(* IEC 61131-3 sources: P26002_Bosch_HDPump/P26002_Bosch_HDPump_PLC/RPM_Profiles, 4 files *)

(* ---- FB_ArrayProfile.st ---- *)
(********************************************************************************
 * FUNCTION_BLOCK: FB_ArrayProfile
 *
 * Beschreibung:
 *   Liest ein 10-ms-Raster Drehzahlprofil aus dem globalen Array aLapData
 *   und interpoliert im 1-ms-Takt stufenlos linear.
 *   Bei Erreichen von nPointsInLap springt der Zeiger auf 0 zurück und
 *   bLapFinished wird für einen Zyklus TRUE.
 ********************************************************************************)
FUNCTION_BLOCK FB_ArrayProfile
VAR_INPUT
    bExecute        : BOOL;
    nPointsInLap    : DINT; (* Tatsächliche Anzahl Punkte im Zyklus *)
END_VAR
VAR_IN_OUT
    aLapDataBuffer  : ARRAY[0..179999] OF REAL; (* Referenz auf das Daten-Array *)
END_VAR
VAR_OUTPUT
    fRpmOut         : REAL;
    bLapFinished    : BOOL;
END_VAR
VAR
    nIndex          : DINT := 0;
    nSubStep1ms     : INT  := 0;
    fCurrentP       : REAL;
    fNextP          : REAL;
    fDeltaPerMs     : REAL;
END_VAR

bLapFinished := FALSE;

(* Plausibilitätsprüfung *)
IF NOT bExecute OR (nPointsInLap <= 1) OR (nPointsInLap > 180000) THEN
    nIndex       := 0;
    nSubStep1ms  := 0;
    fRpmOut      := 0.0;
    RETURN;
END_IF;

(* Alle 10 ms: Neuer Stützwert aus dem Array *)
IF nSubStep1ms = 0 THEN
    fCurrentP := aLapDataBuffer[nIndex];

    (* Nächsten Punkt für Steigungsberechnung holen *)
    IF (nIndex + 1) < nPointsInLap THEN
        fNextP := aLapDataBuffer[nIndex + 1];
    ELSE
        fNextP := aLapDataBuffer[0]; (* Zyklischer Sprung zum Anfang *)
    END_IF;

    (* Steigung pro 1 ms berechnen *)
    fDeltaPerMs := (fNextP - fCurrentP) / 10.0;

    nIndex := nIndex + 1;

    (* RUNDENENDE: Letzter Punkt des Profils erreicht *)
    IF nIndex >= nPointsInLap THEN
        nIndex       := 0;    (* Für nächste Runde zurücksetzen *)
        bLapFinished := TRUE; (* Lap-Signal auslösen *)
    END_IF;
END_IF;

(* 1-ms-Interpolation *)
fRpmOut := fCurrentP + (fDeltaPerMs * INT_TO_REAL(nSubStep1ms));

(* 1-ms-Zähler 0 bis 9 *)
nSubStep1ms := (nSubStep1ms + 1) MOD 10;

END_FUNCTION_BLOCK

(* ---- FB_SequenceController.st ---- *)
(********************************************************************************
 * FUNCTION_BLOCK: FB_SequenceController
 *
 * Beschreibung:
 *   Steuert den Gesamt-Ablauf (Start/Stop, Wiederholungen, Gesamtdauer).
 *   Ausgänge:
 *     - bSequenceActive: TRUE ab Start bis zum Ende der gesamten Sequenz
 *     - bLapTrigger:     Gepulster Ausgang (z.B. 50ms) nach jedem Lap-Durchlauf
 ********************************************************************************)
FUNCTION_BLOCK FB_SequenceController
VAR_INPUT
    bStart              : BOOL;
    bStop               : BOOL;
    eEndMode            : E_SequenceEndMode;
    nTargetLaps         : UDINT;
    tTargetDuration     : TIME;
    tLapPulseDuration   : TIME := T#50ms; (* Einstellbare Pulsdauer *)
    bLapFinishedSignal  : BOOL;
    tCycleTime          : TIME := T#1ms;
END_VAR
VAR_OUTPUT
    bSequenceActive     : BOOL; (* Start/End-Trigger *)
    bLapTrigger         : BOOL; (* Gepulster Lap-Trigger *)
    nCompletedLaps      : UDINT;
    tElapsedTime        : TIME;
END_VAR
VAR
    bStartOld           : BOOL;
    nPulseCyclesLeft    : DINT := 0; (* Exakter Zyklustimer für den Puls *)
END_VAR

(* Stop-Befehl *)
IF bStop THEN
    bSequenceActive  := FALSE;
    nPulseCyclesLeft := 0;
END_IF;

(* Start-Flanke *)
IF bStart AND NOT bStartOld AND NOT bSequenceActive THEN
    bSequenceActive  := TRUE;
    nCompletedLaps   := 0;
    tElapsedTime     := T#0s;
    nPulseCyclesLeft := 0;
END_IF;
bStartOld := bStart;

(* Sequenz-Ablauf *)
IF bSequenceActive THEN
    tElapsedTime := tElapsedTime + tCycleTime;

    (* Lap-Ende registriert *)
    IF bLapFinishedSignal THEN
        nCompletedLaps   := nCompletedLaps + 1;
        (* Millisekunden in 1ms-Taskzyklen konvertieren *)
        nPulseCyclesLeft := TIME_TO_DINT(tLapPulseDuration);
    END_IF;

    (* Abbruchbedingungen *)
    CASE eEndMode OF
        MODE_LAP_COUNT:
            IF nCompletedLaps >= nTargetLaps THEN
                bSequenceActive := FALSE;
            END_IF;

        MODE_TIME_LIMIT:
            IF tElapsedTime >= tTargetDuration THEN
                bSequenceActive := FALSE;
            END_IF;
    END_CASE;
END_IF;

(* Deterministischer Puls über Zyklencounter *)
IF nPulseCyclesLeft > 0 THEN
    bLapTrigger      := TRUE;
    nPulseCyclesLeft := nPulseCyclesLeft - 1;
ELSE
    bLapTrigger := FALSE;
END_IF;

END_FUNCTION_BLOCK

(* ---- FB_SineProfile.st ---- *)
(********************************************************************************
 * FUNCTION_BLOCK: FB_SineProfile
 *
 * Beschreibung:
 *   Erzeugt im 1-ms-Takt ein Sinus-Drehzahlprofil zwischen fRpmMin und fRpmMax
 *   mit parametrierbarer Periodendauer und Phasenversatz in Grad.
 *   Am Ende jeder Periode (tPeriod) wird bLapFinished fuer einen Takt TRUE.
 ********************************************************************************)
FUNCTION_BLOCK FB_SineProfile
VAR_INPUT
    bExecute        : BOOL;
    stConfig        : ST_SineConfig;
    tCycleTime      : TIME := T#1ms;
END_VAR
VAR_OUTPUT
    fRpmOut         : REAL;
    bLapFinished    : BOOL;
END_VAR
VAR
    tCurrentLapTime : TIME := T#0s;
    fOffset         : REAL;
    fAmplitude      : REAL;
    fPeriodSec      : REAL;
    fCurSec         : REAL;
    fPhaseRad       : REAL;
    fAngleRad       : REAL;
END_VAR
VAR CONSTANT
    C_PI            : REAL := 3.14159265;
    C_DEG_TO_RAD    : REAL := 0.0174532925; (* PI / 180.0 *)
END_VAR

bLapFinished := FALSE;

IF NOT bExecute THEN
    tCurrentLapTime := T#0s;
    fRpmOut         := stConfig.fRpmMin;
    RETURN;
END_IF;

fPeriodSec := TIME_TO_REAL(stConfig.tPeriod) / 1000.0;
fCurSec    := TIME_TO_REAL(tCurrentLapTime) / 1000.0;

(* Schutz vor Division durch 0 *)
IF fPeriodSec <= 0.0 THEN
    fRpmOut := stConfig.fRpmMin;
    RETURN;
END_IF;

(* 1. Mittelwert (Offset) und Amplitude berechnen *)
fOffset    := (stConfig.fRpmMax + stConfig.fRpmMin) / 2.0;
fAmplitude := (stConfig.fRpmMax - stConfig.fRpmMin) / 2.0;

(* 2. Phasenversatz und aktuellen Winkel in Bogenmass berechnen *)
fPhaseRad := stConfig.fPhaseDeg * C_DEG_TO_RAD;
fAngleRad := ((2.0 * C_PI / fPeriodSec) * fCurSec) + fPhaseRad;

(* 3. Sollwert ueber Standard-IEC SIN-Funktion berechnen *)
fRpmOut := fOffset + (fAmplitude * SIN(fAngleRad));

(* 4. Zeittakt weiterschalten (1 ms) *)
tCurrentLapTime := tCurrentLapTime + tCycleTime;

(* 5. Periodenende (Lap) erkennen *)
IF tCurrentLapTime >= stConfig.tPeriod THEN
    tCurrentLapTime := T#0s;
    bLapFinished    := TRUE;
END_IF;

END_FUNCTION_BLOCK

(* ---- FB_TriangleProfile.st ---- *)
(********************************************************************************
 * FUNCTION_BLOCK: FB_TriangleProfile
 *
 * Beschreibung:
 *   Erzeugt im 1-ms-Takt ein symmetrisches oder asymmetrisches Dreiecksprofil
 *   zwischen fRpmMin und fRpmMax.
 *   Am Ende der Rampe wird bLapFinished für genau einen Takt TRUE.
 ********************************************************************************)
FUNCTION_BLOCK FB_TriangleProfile
VAR_INPUT
    bExecute        : BOOL;
    stConfig        : ST_TriangleConfig;
    tCycleTime      : TIME := T#1ms;
END_VAR
VAR_OUTPUT
    fRpmOut         : REAL;
    bLapFinished    : BOOL;
END_VAR
VAR
    tCurrentLapTime : TIME := T#0s;
    tRampDownEff    : TIME;
    tTotalLapTime   : TIME;
    fUpSec          : REAL;
    fDownSec        : REAL;
    fCurSec         : REAL;
    fDeltaRpm       : REAL;
END_VAR

bLapFinished := FALSE;

IF NOT bExecute THEN
    tCurrentLapTime := T#0s;
    fRpmOut         := stConfig.fRpmMin;
    RETURN;
END_IF;

(* 1. Symmetrie auswerten *)
IF stConfig.bSymmetric THEN
    tRampDownEff := stConfig.tRampUp;
ELSE
    tRampDownEff := stConfig.tRampDown;
END_IF;

tTotalLapTime := stConfig.tRampUp + tRampDownEff;
fDeltaRpm     := stConfig.fRpmMax - stConfig.fRpmMin;

fUpSec   := TIME_TO_REAL(stConfig.tRampUp) / 1000.0;
fDownSec := TIME_TO_REAL(tRampDownEff) / 1000.0;
fCurSec  := TIME_TO_REAL(tCurrentLapTime) / 1000.0;

(* 2. Rampe berechnen *)
IF tCurrentLapTime < stConfig.tRampUp THEN
    (* Phase 1: Anstieg von Min nach Max *)
    IF fUpSec > 0.0 THEN
        fRpmOut := stConfig.fRpmMin + (fDeltaRpm * (fCurSec / fUpSec));
    ELSE
        fRpmOut := stConfig.fRpmMax;
    END_IF;
ELSE
    (* Phase 2: Abstieg von Max nach Min *)
    IF fDownSec > 0.0 THEN
        fRpmOut := stConfig.fRpmMax - (fDeltaRpm * ((fCurSec - fUpSec) / fDownSec));
    ELSE
        fRpmOut := stConfig.fRpmMin;
    END_IF;
END_IF;

(* 3. Zeittakt weiterschalten (1 ms) *)
tCurrentLapTime := tCurrentLapTime + tCycleTime;

(* 4. Rundenende prüfen *)
IF tCurrentLapTime >= tTotalLapTime THEN
    tCurrentLapTime := T#0s;
    bLapFinished    := TRUE;
END_IF;

END_FUNCTION_BLOCK
